// TIA Portal V20 export
// export: Created 2026-10-19T18:06:26.0866612Z, ExportSetting WithDefaults, DisplayName Totally Integrated Automation Portal, DisplayVersion V20 Update 6, DisplayName TIA Portal Openness, DisplayVersion V20 Update 6, DisplayName TIA Portal Version Control Interface, DisplayVersion V20 Update 6, DisplayName SINAMICS Startdrive Advanced, DisplayVersion V20 SP1, DisplayName SINAMICS Startdrive G130, G150, S120, S150, SINAMICS MV, G220, S200, S210, DisplayVersion V20 SP1, DisplayName SINAMICS Startdrive G110M, G120, G120C, G120D, G120P, G115D, DisplayVersion V20 SP1, DisplayName STEP 7 Professional, DisplayVersion V20 Update 6, DisplayName STEP 7 Safety, DisplayVersion V20 Update 2, DisplayName WinCC Basic/Comfort/Advanced, DisplayVersion V20 Update 6, DisplayName WinCC Unified, DisplayVersion V20 Update 6
FUNCTION_BLOCK "SAI_IND_SpanAdjust"   // FB55, LAD
TITLE = Span and Linearity Adjustment (Multi-Point Selectable)
{ S7_Optimized_Access := 'FALSE' }
VERSION : 0.1
// stored: AutoNumber true, IsIECCheckEnabled false, SetENOAutomatically false, UDAEnableTagReadback false
   VAR_INPUT
      ID : HW_IO;   // The Profinet Device Hardware Identifier under device properties
      Hi_Weight : Real;   // The highest adjustment weight, or the Span value
      Mid_Weight : Real;   // The 4th adjustment weight
      Low_Weight : Real;   // The 3rd adjustment weight
      xLow_Weight : Real;   // The 2nd adjustment weight
   END_VAR
   VAR_OUTPUT
      CurrentPoint : Int;   // Current point to be adjusted (Minimum 2 points; maximum 5 points; zero point is the 1st point)
      CurrentWeight : Real;   // Current adjustment weight to be loaded onto the scale
      LoadWeight : Bool;   // Load the next adjustment weight according to value shown in CurrentWeight
      Process : Bool;   // Weight Transmitter is performing adjustment
      Done : Bool;   // Linearity Adjustment has been completed successfully
      Error : Bool;   // Adjustment can not proceed due to incomplete input parameters, check LinearityRange and all the adjustment weight values
      Cancelled : Bool;   // Adjustment process has been cancelled successfully
   END_VAR
   VAR_IN_OUT
      LinearityRange : Int;   // Number of linearity points to be adjusted: 0:none, 1:3 point, 2:4 point, 3:5 point
      Start : Bool;   // Trigger this bit ON to start performing linearity adjustment; this bit will be turned off automatically after completion
      ConfirmWeight : Bool;   // Switch ON this bit as an acknowledgement that new adjustment weight has being loaded
      Cancel : Bool;   // Cancel/ Abort adjustment process, toggle ON
   END_VAR
   VAR DB_SPECIFIC
      Activate : Bool;
   END_VAR
   VAR
      WRREC_SpanAdjust { S7_SetPoint := 'True'} : WRREC;
      RDREC_Status { S7_SetPoint := 'True'} : RDREC;
   END_VAR
   VAR DB_SPECIFIC
      IEC_Timer_1_Instance { S7_SetPoint := 'True'} : IEC_TIMER;
      AdjustStep : SInt;
      Static01 : Bool;
      Static02 : Bool;
      Static03 : Bool;
      Static04 : Bool;
      Static05 : Bool;
      Static06 : Bool;
      Static07 : Bool;
      Static08 : Bool;
      Validate_REC : SInt;
      Abort_REC : SInt;
      Check01 : Bool;
      Check02 : Bool;
      AdjustmentStatus : Int;
      CurrentPoint_0 : Int;
      CurrentWeight_0 : Real;
   END_VAR
   VAR_TEMP   // added for the SCL form of the ladder/FBD networks
      _w1 : Bool;
      _w2 : Bool;
      _w3 : Bool;
      _w4 : Bool;
      _w5 : Bool;
      _w6 : Bool;
      _w7 : Bool;
      _w8 : Bool;
      _w9 : Bool;
      _w10 : Bool;
      _w11 : Bool;
      _w12 : Bool;
      _w13 : Bool;
   END_VAR
BEGIN

REGION Network 1: Initialization
   // Initializes FB output bits:
   // Process;
   // Error;
   // Done;
   // Cancelled
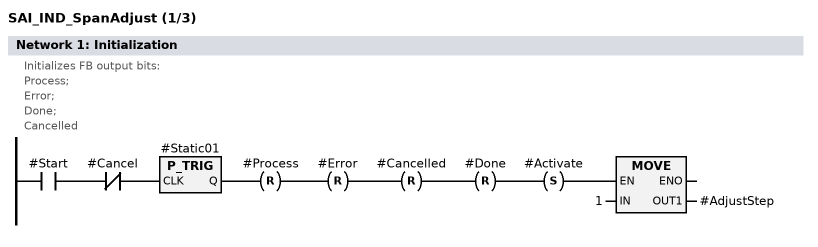
   RUNG wire#powerrail
      Contact( #Start )
      I_Contact( #Cancel )
      P_Trig( #Static01 )
      R_Coil( #Process )
      R_Coil( #Error )
      R_Coil( #Cancelled )
      R_Coil( #Done )
      S_Coil( #Activate )
      { S7_GenerateENO := "TRUE" } Move(in := 1, out1 => #AdjustStep)
   END_RUNG
   // the same network as SCL:
   #_w1 := #Start AND NOT #Cancel;
   #_w2 := #_w1 AND NOT #Static01;   // rising edge
   #Static01 := #_w1;
   IF #_w2 THEN
       #Process := FALSE;
       #Error := FALSE;
       #Cancelled := FALSE;
       #Done := FALSE;
       #Activate := TRUE;
       #AdjustStep := 1;
   END_IF;
END_REGION

REGION Network 2: Sequence
   // AdjustStep = 1: Check all the input parameters for LinearityRange and adjustment weights (Hi_Weight, Mid_Weight, Low_Weight, xLow_Weight)
   // AdjustStep = 2: Initializes all the control bits
   // AdjustStep = 3: Write in the LinearityRange into the transmitter (2-byte; Index: 16#400A)
   // AdjustStep = 4: Updates the CurrentPoint and CurrentWeight (new reference weight) and wait for user to trigger ConfirmWeight input bit
   // AdjustStep = 5: Start the adjustment process according to the CurrentWeight (REAL; Index: 16#4009)
   // AdjustStep = 6: After adjusted all the required reference weights, validate the adjustment (2-byte; Index: 16#4010)
   // AdjustStep = 7: Adjustment is completed successfully, set DONE bit to TRUE
   // AdjustStep = 8; Adjustment failed with error, set ERROR bit to TRUE
   // AdjustStep >= 4: Reading the adjustment status continuously (2-byte; Index: 16#4007)
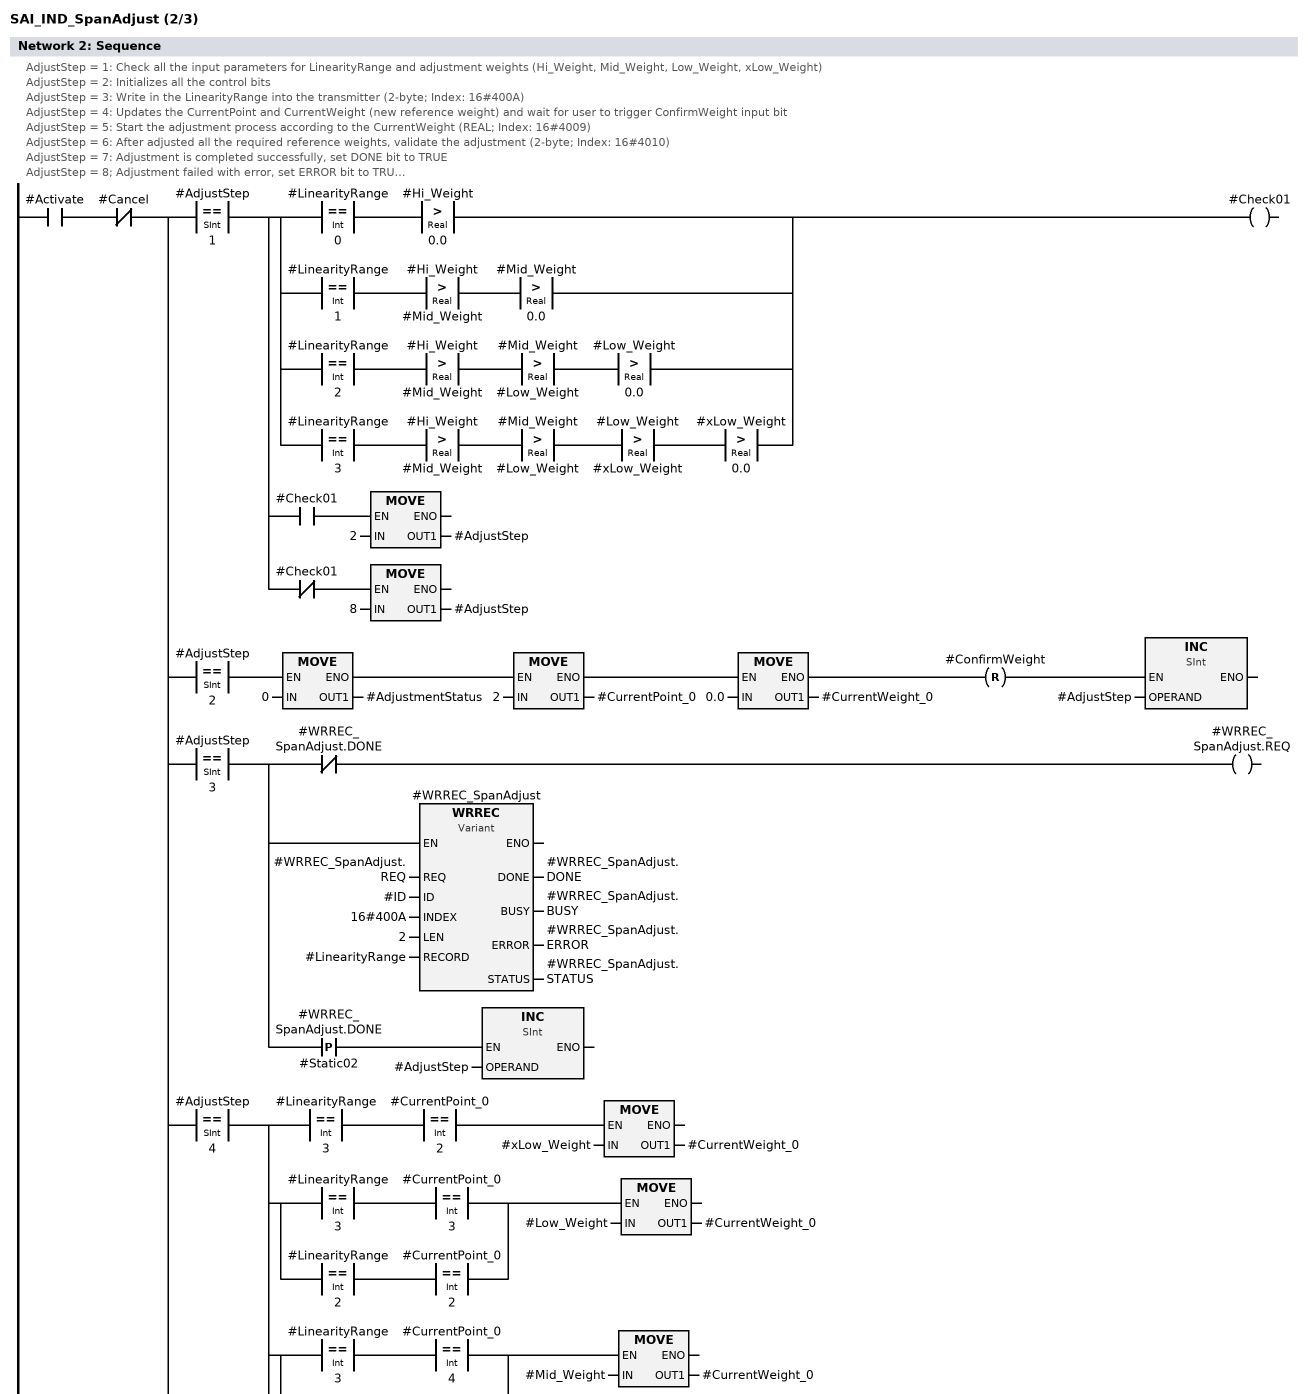
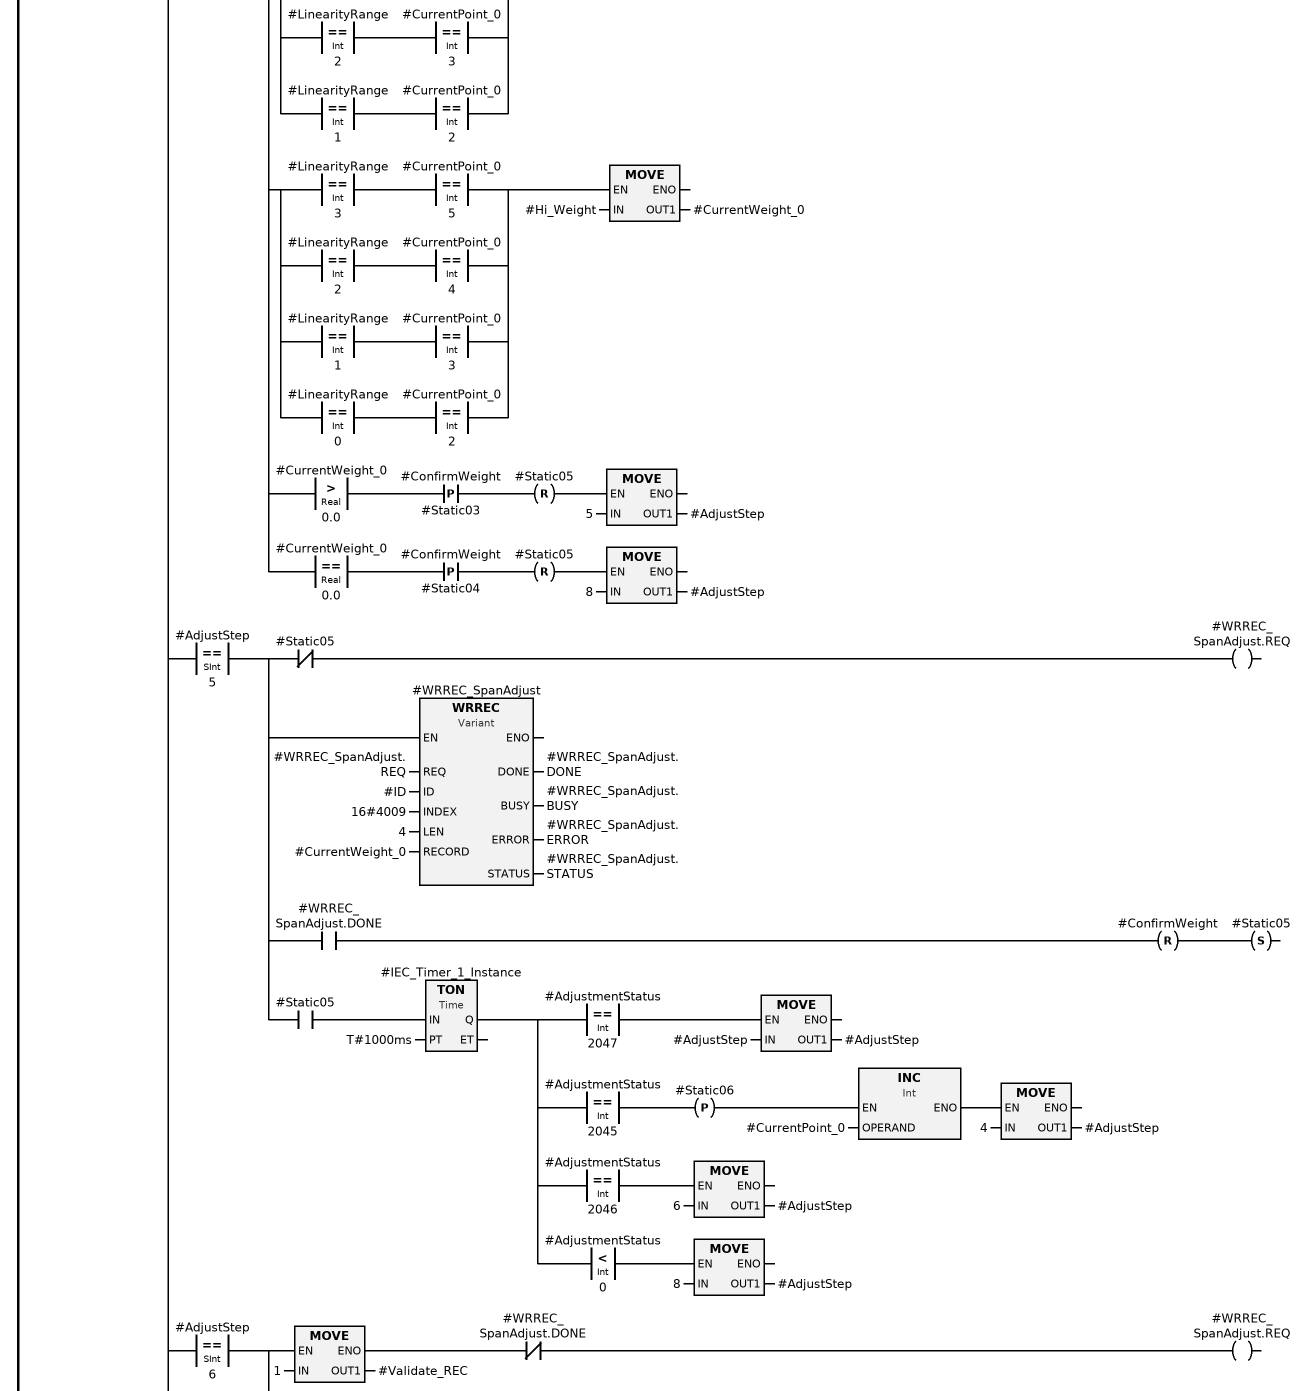
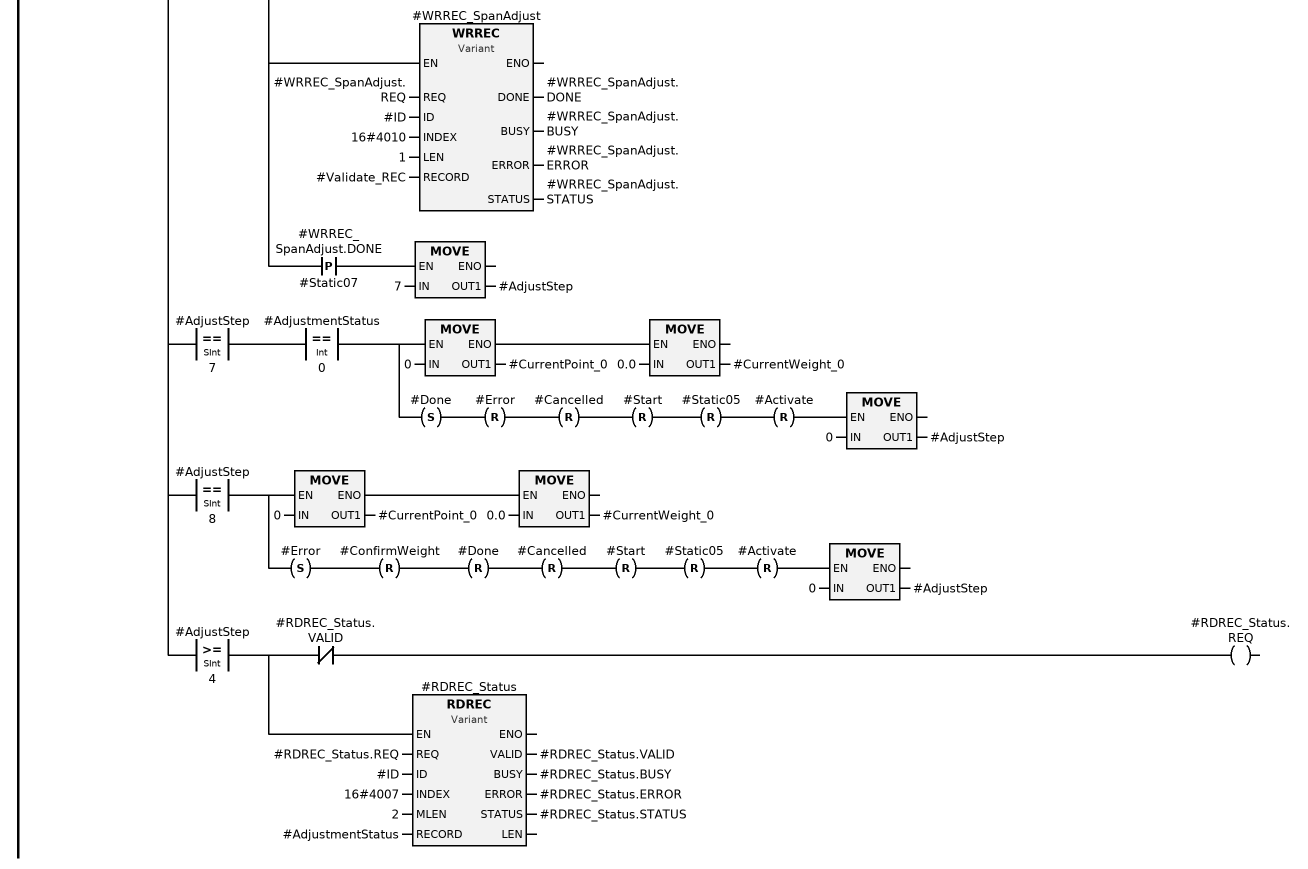
   RUNG wire#powerrail
      Contact( #Activate )
      I_Contact( #Cancel )
      wire#w1
      { S7_Templates := "SrcType := SInt" } EQ_Contact(in1 := #AdjustStep, in2 := 1)
      wire#w2
      { S7_Templates := "SrcType := Int" } EQ_Contact(in1 := #LinearityRange, in2 := 0)
      { S7_Templates := "SrcType := Real" } GT_Contact(in1 := #Hi_Weight, in2 := 0.0)
      wire#w3
      Coil( #Check01 )
   END_RUNG
   RUNG wire#w2
      { S7_Templates := "SrcType := Int" } EQ_Contact(in1 := #LinearityRange, in2 := 1)
      { S7_Templates := "SrcType := Real" } GT_Contact(in1 := #Hi_Weight, in2 := #Mid_Weight)
      { S7_Templates := "SrcType := Real" } GT_Contact(in1 := #Mid_Weight, in2 := 0.0)
   END_RUNG wire#w3
   RUNG wire#w2
      { S7_Templates := "SrcType := Int" } EQ_Contact(in1 := #LinearityRange, in2 := 2)
      { S7_Templates := "SrcType := Real" } GT_Contact(in1 := #Hi_Weight, in2 := #Mid_Weight)
      { S7_Templates := "SrcType := Real" } GT_Contact(in1 := #Mid_Weight, in2 := #Low_Weight)
      { S7_Templates := "SrcType := Real" } GT_Contact(in1 := #Low_Weight, in2 := 0.0)
   END_RUNG wire#w3
   RUNG wire#w2
      { S7_Templates := "SrcType := Int" } EQ_Contact(in1 := #LinearityRange, in2 := 3)
      { S7_Templates := "SrcType := Real" } GT_Contact(in1 := #Hi_Weight, in2 := #Mid_Weight)
      { S7_Templates := "SrcType := Real" } GT_Contact(in1 := #Mid_Weight, in2 := #Low_Weight)
      { S7_Templates := "SrcType := Real" } GT_Contact(in1 := #Low_Weight, in2 := #xLow_Weight)
      { S7_Templates := "SrcType := Real" } GT_Contact(in1 := #xLow_Weight, in2 := 0.0)
   END_RUNG wire#w3
   RUNG wire#w2
      Contact( #Check01 )
      Move(in := 2, out1 => #AdjustStep)
   END_RUNG
   RUNG wire#w2
      I_Contact( #Check01 )
      Move(in := 8, out1 => #AdjustStep)
   END_RUNG
   RUNG wire#w1
      { S7_Templates := "SrcType := SInt" } EQ_Contact(in1 := #AdjustStep, in2 := 2)
      Move(in := 0, out1 => #AdjustmentStatus)
      Move(in := 2, out1 => #CurrentPoint_0)
      Move(in := 0.0, out1 => #CurrentWeight_0)
      R_Coil( #ConfirmWeight )
      { S7_Templates := "DestType := SInt" } Inc( #AdjustStep )
   END_RUNG
   RUNG wire#w1
      { S7_Templates := "SrcType := SInt" } EQ_Contact(in1 := #AdjustStep, in2 := 3)
      wire#w4
      I_Contact( #WRREC_SpanAdjust.DONE )
      Coil( #WRREC_SpanAdjust.REQ )
   END_RUNG
   RUNG wire#w4
      { S7_Templates := "[ptr_type := Variant, id_type := HW_IO, index_type := DInt, len_type := UInt]" } #WRREC_SpanAdjust.WRREC(REQ := #WRREC_SpanAdjust.REQ, ID := #ID, INDEX := 16#400A, LEN := 2, RECORD := #LinearityRange, DONE => #WRREC_SpanAdjust.DONE, BUSY => #WRREC_SpanAdjust.BUSY, ERROR => #WRREC_SpanAdjust.ERROR, STATUS => #WRREC_SpanAdjust.STATUS)
   END_RUNG
   RUNG wire#w4
      P_Contact(operand := #WRREC_SpanAdjust.DONE, bit := #Static02)
      { S7_Templates := "DestType := SInt" } Inc( #AdjustStep )
   END_RUNG
   RUNG wire#w1
      { S7_Templates := "SrcType := SInt" } EQ_Contact(in1 := #AdjustStep, in2 := 4)
      wire#w5
      { S7_Templates := "SrcType := Int" } EQ_Contact(in1 := #LinearityRange, in2 := 3)
      { S7_Templates := "SrcType := Int" } EQ_Contact(in1 := #CurrentPoint_0, in2 := 2)
      Move(in := #xLow_Weight, out1 => #CurrentWeight_0)
   END_RUNG
   RUNG wire#w5
      { S7_Templates := "SrcType := Int" } EQ_Contact(in1 := #LinearityRange, in2 := 3)
      { S7_Templates := "SrcType := Int" } EQ_Contact(in1 := #CurrentPoint_0, in2 := 3)
      wire#w6
      Move(in := #Low_Weight, out1 => #CurrentWeight_0)
   END_RUNG
   RUNG wire#w5
      { S7_Templates := "SrcType := Int" } EQ_Contact(in1 := #LinearityRange, in2 := 2)
      { S7_Templates := "SrcType := Int" } EQ_Contact(in1 := #CurrentPoint_0, in2 := 2)
   END_RUNG wire#w6
   RUNG wire#w5
      { S7_Templates := "SrcType := Int" } EQ_Contact(in1 := #LinearityRange, in2 := 3)
      { S7_Templates := "SrcType := Int" } EQ_Contact(in1 := #CurrentPoint_0, in2 := 4)
      wire#w7
      Move(in := #Mid_Weight, out1 => #CurrentWeight_0)
   END_RUNG
   RUNG wire#w5
      { S7_Templates := "SrcType := Int" } EQ_Contact(in1 := #LinearityRange, in2 := 2)
      { S7_Templates := "SrcType := Int" } EQ_Contact(in1 := #CurrentPoint_0, in2 := 3)
   END_RUNG wire#w7
   RUNG wire#w5
      { S7_Templates := "SrcType := Int" } EQ_Contact(in1 := #LinearityRange, in2 := 1)
      { S7_Templates := "SrcType := Int" } EQ_Contact(in1 := #CurrentPoint_0, in2 := 2)
   END_RUNG wire#w7
   RUNG wire#w5
      { S7_Templates := "SrcType := Int" } EQ_Contact(in1 := #LinearityRange, in2 := 3)
      { S7_Templates := "SrcType := Int" } EQ_Contact(in1 := #CurrentPoint_0, in2 := 5)
      wire#w8
      Move(in := #Hi_Weight, out1 => #CurrentWeight_0)
   END_RUNG
   RUNG wire#w5
      { S7_Templates := "SrcType := Int" } EQ_Contact(in1 := #LinearityRange, in2 := 2)
      { S7_Templates := "SrcType := Int" } EQ_Contact(in1 := #CurrentPoint_0, in2 := 4)
   END_RUNG wire#w8
   RUNG wire#w5
      { S7_Templates := "SrcType := Int" } EQ_Contact(in1 := #LinearityRange, in2 := 1)
      { S7_Templates := "SrcType := Int" } EQ_Contact(in1 := #CurrentPoint_0, in2 := 3)
   END_RUNG wire#w8
   RUNG wire#w5
      { S7_Templates := "SrcType := Int" } EQ_Contact(in1 := #LinearityRange, in2 := 0)
      { S7_Templates := "SrcType := Int" } EQ_Contact(in1 := #CurrentPoint_0, in2 := 2)
   END_RUNG wire#w8
   RUNG wire#w5
      { S7_Templates := "SrcType := Real" } GT_Contact(in1 := #CurrentWeight_0, in2 := 0.0)
      P_Contact(operand := #ConfirmWeight, bit := #Static03)
      R_Coil( #Static05 )
      Move(in := 5, out1 => #AdjustStep)
   END_RUNG
   RUNG wire#w5
      { S7_Templates := "SrcType := Real" } EQ_Contact(in1 := #CurrentWeight_0, in2 := 0.0)
      P_Contact(operand := #ConfirmWeight, bit := #Static04)
      R_Coil( #Static05 )
      Move(in := 8, out1 => #AdjustStep)
   END_RUNG
   RUNG wire#w1
      { S7_Templates := "SrcType := SInt" } EQ_Contact(in1 := #AdjustStep, in2 := 5)
      wire#w9
      I_Contact( #Static05 )
      Coil( #WRREC_SpanAdjust.REQ )
   END_RUNG
   RUNG wire#w9
      { S7_Templates := "[ptr_type := Variant, id_type := HW_IO, index_type := DInt, len_type := UInt]" } #WRREC_SpanAdjust.WRREC(REQ := #WRREC_SpanAdjust.REQ, ID := #ID, INDEX := 16#4009, LEN := 4, RECORD := #CurrentWeight_0, DONE => #WRREC_SpanAdjust.DONE, BUSY => #WRREC_SpanAdjust.BUSY, ERROR => #WRREC_SpanAdjust.ERROR, STATUS => #WRREC_SpanAdjust.STATUS)
   END_RUNG
   RUNG wire#w9
      Contact( #WRREC_SpanAdjust.DONE )
      R_Coil( #ConfirmWeight )
      S_Coil( #Static05 )
   END_RUNG
   RUNG wire#w9
      Contact( #Static05 )
      { S7_Templates := "time_type := Time" } #IEC_Timer_1_Instance.TON(pt := T#1000ms, et =>)
      wire#w10
      { S7_Templates := "SrcType := Int" } EQ_Contact(in1 := #AdjustmentStatus, in2 := 2047)
      Move(in := #AdjustStep, out1 => #AdjustStep)
   END_RUNG
   RUNG wire#w10
      { S7_Templates := "SrcType := Int" } EQ_Contact(in1 := #AdjustmentStatus, in2 := 2045)
      P_Trig( #Static06 )
      { S7_Templates := "DestType := Int" } Inc( #CurrentPoint_0 )
      Move(in := 4, out1 => #AdjustStep)
   END_RUNG
   RUNG wire#w10
      { S7_Templates := "SrcType := Int" } EQ_Contact(in1 := #AdjustmentStatus, in2 := 2046)
      Move(in := 6, out1 => #AdjustStep)
   END_RUNG
   RUNG wire#w10
      { S7_Templates := "SrcType := Int" } LT_Contact(in1 := #AdjustmentStatus, in2 := 0)
      Move(in := 8, out1 => #AdjustStep)
   END_RUNG
   RUNG wire#w1
      { S7_Templates := "SrcType := SInt" } EQ_Contact(in1 := #AdjustStep, in2 := 6)
      wire#w11
      Move(in := 1, out1 => #Validate_REC)
      I_Contact( #WRREC_SpanAdjust.DONE )
      Coil( #WRREC_SpanAdjust.REQ )
   END_RUNG
   RUNG wire#w11
      { S7_Templates := "[ptr_type := Variant, id_type := HW_IO, index_type := DInt, len_type := UInt]" } #WRREC_SpanAdjust.WRREC(REQ := #WRREC_SpanAdjust.REQ, ID := #ID, INDEX := 16#4010, LEN := 1, RECORD := #Validate_REC, DONE => #WRREC_SpanAdjust.DONE, BUSY => #WRREC_SpanAdjust.BUSY, ERROR => #WRREC_SpanAdjust.ERROR, STATUS => #WRREC_SpanAdjust.STATUS)
   END_RUNG
   RUNG wire#w11
      P_Contact(operand := #WRREC_SpanAdjust.DONE, bit := #Static07)
      Move(in := 7, out1 => #AdjustStep)
   END_RUNG
   RUNG wire#w1
      { S7_Templates := "SrcType := SInt" } EQ_Contact(in1 := #AdjustStep, in2 := 7)
      { S7_Templates := "SrcType := Int" } EQ_Contact(in1 := #AdjustmentStatus, in2 := 0)
      wire#w12
      Move(in := 0, out1 => #CurrentPoint_0)
      Move(in := 0.0, out1 => #CurrentWeight_0)
   END_RUNG
   RUNG wire#w12
      S_Coil( #Done )
      R_Coil( #Error )
      R_Coil( #Cancelled )
      R_Coil( #Start )
      R_Coil( #Static05 )
      R_Coil( #Activate )
      Move(in := 0, out1 => #AdjustStep)
   END_RUNG
   RUNG wire#w1
      { S7_Templates := "SrcType := SInt" } EQ_Contact(in1 := #AdjustStep, in2 := 8)
      wire#w13
      Move(in := 0, out1 => #CurrentPoint_0)
      Move(in := 0.0, out1 => #CurrentWeight_0)
   END_RUNG
   RUNG wire#w13
      S_Coil( #Error )
      R_Coil( #ConfirmWeight )
      R_Coil( #Done )
      R_Coil( #Cancelled )
      R_Coil( #Start )
      R_Coil( #Static05 )
      R_Coil( #Activate )
      Move(in := 0, out1 => #AdjustStep)
   END_RUNG
   RUNG wire#w1
      { S7_Templates := "SrcType := SInt" } GE_Contact(in1 := #AdjustStep, in2 := 4)
      wire#w14
      I_Contact( #RDREC_Status.VALID )
      Coil( #RDREC_Status.REQ )
   END_RUNG
   RUNG wire#w14
      { S7_Templates := "[ptr_type := Variant, id_type := HW_IO, index_type := DInt, len_type := UInt]" } #RDREC_Status.RDREC(REQ := #RDREC_Status.REQ, ID := #ID, INDEX := 16#4007, MLEN := 2, RECORD := #AdjustmentStatus, VALID => #RDREC_Status.VALID, BUSY => #RDREC_Status.BUSY, ERROR => #RDREC_Status.ERROR, STATUS => #RDREC_Status.STATUS, LEN =>)
   END_RUNG
   // the same network as SCL:
   #_w1 := #Activate AND NOT #Cancel;
   #_w2 := #_w1 AND (#AdjustStep = 1);
   #Check01 := #_w2 AND (((#LinearityRange = 0) AND (#Hi_Weight > 0.0)) OR ((#LinearityRange = 1) AND (#Hi_Weight > #Mid_Weight) AND (#Mid_Weight > 0.0)) OR ((#LinearityRange = 2) AND (#Hi_Weight > #Mid_Weight) AND (#Mid_Weight > #Low_Weight) AND (#Low_Weight > 0.0)) OR ((#LinearityRange = 3) AND (#Hi_Weight > #Mid_Weight) AND (#Mid_Weight > #Low_Weight) AND (#Low_Weight > #xLow_Weight) AND (#xLow_Weight > 0.0)));
   IF #_w2 AND #Check01 THEN #AdjustStep := 2; END_IF;
   IF #_w2 AND NOT #Check01 THEN #AdjustStep := 8; END_IF;
   IF #_w1 AND (#AdjustStep = 2) THEN
       #AdjustmentStatus := 0;
       #CurrentPoint_0 := 2;
       #CurrentWeight_0 := 0.0;
       #ConfirmWeight := FALSE;
       #AdjustStep := #AdjustStep + 1;
   END_IF;
   #_w3 := #_w1 AND (#AdjustStep = 3);
   #WRREC_SpanAdjust.REQ := #_w3 AND NOT #WRREC_SpanAdjust.DONE;
   IF #_w3 THEN
       #WRREC_SpanAdjust(REQ := #WRREC_SpanAdjust.REQ,   // WRREC
                         ID := #ID,
                         INDEX := 16#400A,
                         LEN := 2,
                         RECORD := #LinearityRange,
                         DONE => #WRREC_SpanAdjust.DONE,
                         BUSY => #WRREC_SpanAdjust.BUSY,
                         ERROR => #WRREC_SpanAdjust.ERROR,
                         STATUS => #WRREC_SpanAdjust.STATUS);
   END_IF;
   #_w4 := #_w3 AND #WRREC_SpanAdjust.DONE AND NOT #Static02;   // rising edge of #WRREC_SpanAdjust.DONE
   #Static02 := #WRREC_SpanAdjust.DONE;
   IF #_w4 THEN #AdjustStep := #AdjustStep + 1; END_IF;
   #_w5 := #_w1 AND (#AdjustStep = 4);
   IF #_w5 AND (#LinearityRange = 3) AND (#CurrentPoint_0 = 2) THEN #CurrentWeight_0 := #xLow_Weight; END_IF;
   IF #_w5 AND (((#LinearityRange = 3) AND (#CurrentPoint_0 = 3)) OR ((#LinearityRange = 2) AND (#CurrentPoint_0 = 2))) THEN
       #CurrentWeight_0 := #Low_Weight;
   END_IF;
   IF #_w5 AND (((#LinearityRange = 3) AND (#CurrentPoint_0 = 4)) OR ((#LinearityRange = 2) AND (#CurrentPoint_0 = 3)) OR ((#LinearityRange = 1) AND (#CurrentPoint_0 = 2))) THEN
       #CurrentWeight_0 := #Mid_Weight;
   END_IF;
   IF #_w5 AND (((#LinearityRange = 3) AND (#CurrentPoint_0 = 5)) OR ((#LinearityRange = 2) AND (#CurrentPoint_0 = 4)) OR ((#LinearityRange = 1) AND (#CurrentPoint_0 = 3)) OR ((#LinearityRange = 0) AND (#CurrentPoint_0 = 2))) THEN
       #CurrentWeight_0 := #Hi_Weight;
   END_IF;
   #_w6 := #_w5 AND (#CurrentWeight_0 > 0.0) AND #ConfirmWeight AND NOT #Static03;   // rising edge of #ConfirmWeight
   #Static03 := #ConfirmWeight;
   IF #_w6 THEN
       #Static05 := FALSE;
       #AdjustStep := 5;
   END_IF;
   #_w7 := #_w5 AND (#CurrentWeight_0 = 0.0) AND #ConfirmWeight AND NOT #Static04;   // rising edge of #ConfirmWeight
   #Static04 := #ConfirmWeight;
   IF #_w7 THEN
       #Static05 := FALSE;
       #AdjustStep := 8;
   END_IF;
   #_w8 := #_w1 AND (#AdjustStep = 5);
   #WRREC_SpanAdjust.REQ := #_w8 AND NOT #Static05;
   IF #_w8 THEN
       #WRREC_SpanAdjust(REQ := #WRREC_SpanAdjust.REQ,   // WRREC
                         ID := #ID,
                         INDEX := 16#4009,
                         LEN := 4,
                         RECORD := #CurrentWeight_0,
                         DONE => #WRREC_SpanAdjust.DONE,
                         BUSY => #WRREC_SpanAdjust.BUSY,
                         ERROR => #WRREC_SpanAdjust.ERROR,
                         STATUS => #WRREC_SpanAdjust.STATUS);
   END_IF;
   IF #_w8 AND #WRREC_SpanAdjust.DONE THEN
       #ConfirmWeight := FALSE;
       #Static05 := TRUE;
   END_IF;
   #IEC_Timer_1_Instance.TON(IN := #_w8 AND #Static05, PT := T#1000ms);
   IF #IEC_Timer_1_Instance.Q AND (#AdjustmentStatus = 2047) THEN #AdjustStep := #AdjustStep; END_IF;
   #_w9 := #IEC_Timer_1_Instance.Q AND (#AdjustmentStatus = 2045);
   #_w10 := #_w9 AND NOT #Static06;   // rising edge
   #Static06 := #_w9;
   IF #_w10 THEN
       #CurrentPoint_0 := #CurrentPoint_0 + 1;
       #AdjustStep := 4;
   END_IF;
   IF #IEC_Timer_1_Instance.Q AND (#AdjustmentStatus = 2046) THEN #AdjustStep := 6; END_IF;
   IF #IEC_Timer_1_Instance.Q AND (#AdjustmentStatus < 0) THEN #AdjustStep := 8; END_IF;
   #_w11 := #_w1 AND (#AdjustStep = 6);
   IF #_w11 THEN #Validate_REC := 1; END_IF;
   #WRREC_SpanAdjust.REQ := #_w11 AND NOT #WRREC_SpanAdjust.DONE;
   IF #_w11 THEN
       #WRREC_SpanAdjust(REQ := #WRREC_SpanAdjust.REQ,   // WRREC
                         ID := #ID,
                         INDEX := 16#4010,
                         LEN := 1,
                         RECORD := #Validate_REC,
                         DONE => #WRREC_SpanAdjust.DONE,
                         BUSY => #WRREC_SpanAdjust.BUSY,
                         ERROR => #WRREC_SpanAdjust.ERROR,
                         STATUS => #WRREC_SpanAdjust.STATUS);
   END_IF;
   #_w12 := #_w11 AND #WRREC_SpanAdjust.DONE AND NOT #Static07;   // rising edge of #WRREC_SpanAdjust.DONE
   #Static07 := #WRREC_SpanAdjust.DONE;
   IF #_w12 THEN #AdjustStep := 7; END_IF;
   IF #_w1 AND (#AdjustStep = 7) AND (#AdjustmentStatus = 0) THEN
       #CurrentPoint_0 := 0;
       #CurrentWeight_0 := 0.0;
       #Done := TRUE;
       #Error := FALSE;
       #Cancelled := FALSE;
       #Start := FALSE;
       #Static05 := FALSE;
       #Activate := FALSE;
       #AdjustStep := 0;
   END_IF;
   IF #_w1 AND (#AdjustStep = 8) THEN
       #CurrentPoint_0 := 0;
       #CurrentWeight_0 := 0.0;
       #Error := TRUE;
       #ConfirmWeight := FALSE;
       #Done := FALSE;
       #Cancelled := FALSE;
       #Start := FALSE;
       #Static05 := FALSE;
       #Activate := FALSE;
       #AdjustStep := 0;
   END_IF;
   #_w13 := #_w1 AND (#AdjustStep >= 4);
   #RDREC_Status.REQ := #_w13 AND NOT #RDREC_Status.VALID;
   IF #_w13 THEN
       #RDREC_Status(REQ := #RDREC_Status.REQ,   // RDREC
                     ID := #ID,
                     INDEX := 16#4007,
                     MLEN := 2,
                     RECORD := #AdjustmentStatus,
                     VALID => #RDREC_Status.VALID,
                     BUSY => #RDREC_Status.BUSY,
                     ERROR => #RDREC_Status.ERROR,
                     STATUS => #RDREC_Status.STATUS);
   END_IF;
END_REGION

REGION Network 3: Adjsutment Status
   // LoadWeight - Inform user to load the next adjustment weight according to CurrentWeight value
   // Process - Status bit to inform that the weight transmitter is performing adjustment process
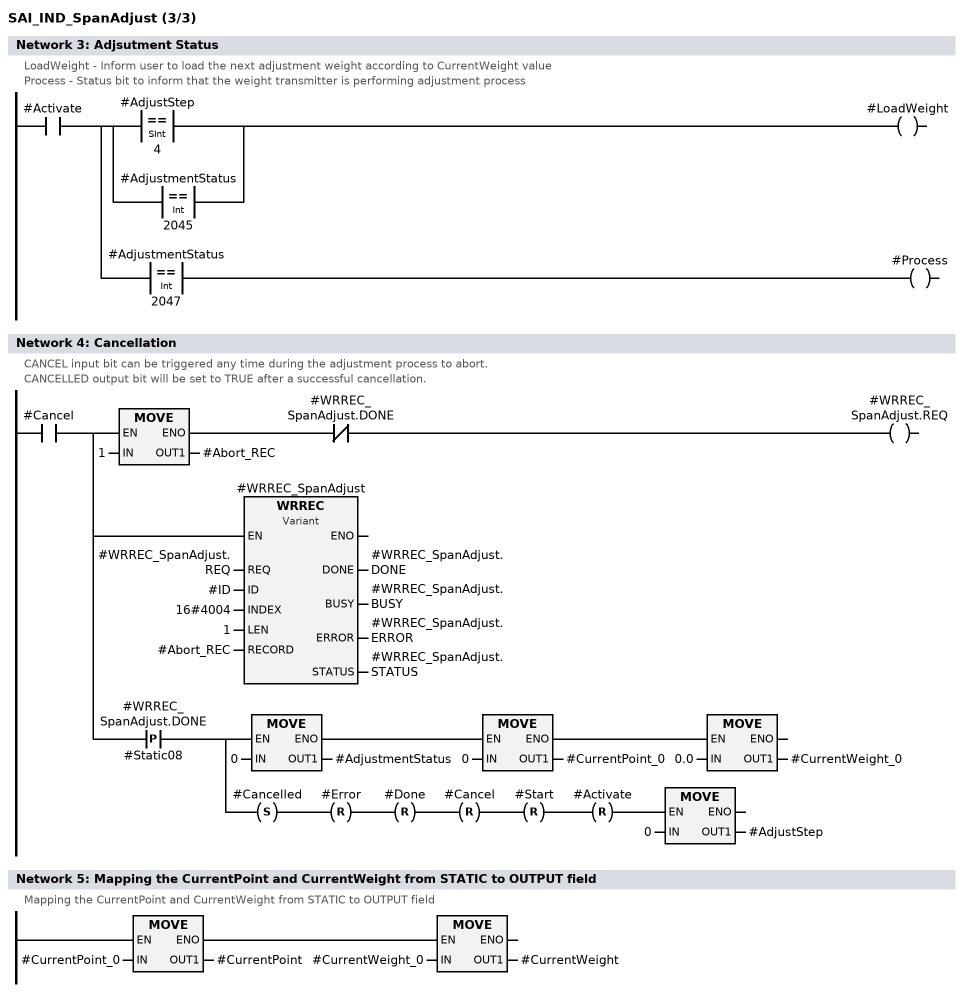
   RUNG wire#powerrail
      Contact( #Activate )
      wire#w1
      { S7_Templates := "SrcType := SInt" } EQ_Contact(in1 := #AdjustStep, in2 := 4)
      wire#w2
      Coil( #LoadWeight )
   END_RUNG
   RUNG wire#w1
      { S7_Templates := "SrcType := Int" } EQ_Contact(in1 := #AdjustmentStatus, in2 := 2045)
   END_RUNG wire#w2
   RUNG wire#w1
      { S7_Templates := "SrcType := Int" } EQ_Contact(in1 := #AdjustmentStatus, in2 := 2047)
      Coil( #Process )
   END_RUNG
   // the same network as SCL:
   #LoadWeight := #Activate AND ((#AdjustStep = 4) OR (#AdjustmentStatus = 2045));
   #Process := #Activate AND (#AdjustmentStatus = 2047);
END_REGION

REGION Network 4: Cancellation
   // CANCEL input bit can be triggered any time during the adjustment process to abort. 
   // CANCELLED output bit will be set to TRUE after a successful cancellation.
   RUNG wire#powerrail
      Contact( #Cancel )
      wire#w1
      Move(in := 1, out1 => #Abort_REC)
      I_Contact( #WRREC_SpanAdjust.DONE )
      Coil( #WRREC_SpanAdjust.REQ )
   END_RUNG
   RUNG wire#w1
      { S7_Templates := "[ptr_type := Variant, id_type := HW_IO, index_type := DInt, len_type := UInt]" } #WRREC_SpanAdjust.WRREC(REQ := #WRREC_SpanAdjust.REQ, ID := #ID, INDEX := 16#4004, LEN := 1, RECORD := #Abort_REC, DONE => #WRREC_SpanAdjust.DONE, BUSY => #WRREC_SpanAdjust.BUSY, ERROR => #WRREC_SpanAdjust.ERROR, STATUS => #WRREC_SpanAdjust.STATUS)
   END_RUNG
   RUNG wire#w1
      P_Contact(operand := #WRREC_SpanAdjust.DONE, bit := #Static08)
      wire#w2
      Move(in := 0, out1 => #AdjustmentStatus)
      Move(in := 0, out1 => #CurrentPoint_0)
      Move(in := 0.0, out1 => #CurrentWeight_0)
   END_RUNG
   RUNG wire#w2
      S_Coil( #Cancelled )
      R_Coil( #Error )
      R_Coil( #Done )
      R_Coil( #Cancel )
      R_Coil( #Start )
      R_Coil( #Activate )
      Move(in := 0, out1 => #AdjustStep)
   END_RUNG
   // the same network as SCL:
   IF #Cancel THEN #Abort_REC := 1; END_IF;
   #WRREC_SpanAdjust.REQ := #Cancel AND NOT #WRREC_SpanAdjust.DONE;
   IF #Cancel THEN
       #WRREC_SpanAdjust(REQ := #WRREC_SpanAdjust.REQ,   // WRREC
                         ID := #ID,
                         INDEX := 16#4004,
                         LEN := 1,
                         RECORD := #Abort_REC,
                         DONE => #WRREC_SpanAdjust.DONE,
                         BUSY => #WRREC_SpanAdjust.BUSY,
                         ERROR => #WRREC_SpanAdjust.ERROR,
                         STATUS => #WRREC_SpanAdjust.STATUS);
   END_IF;
   #_w1 := #Cancel AND #WRREC_SpanAdjust.DONE AND NOT #Static08;   // rising edge of #WRREC_SpanAdjust.DONE
   #Static08 := #WRREC_SpanAdjust.DONE;
   IF #_w1 THEN
       #AdjustmentStatus := 0;
       #CurrentPoint_0 := 0;
       #CurrentWeight_0 := 0.0;
       #Cancelled := TRUE;
       #Error := FALSE;
       #Done := FALSE;
       #Cancel := FALSE;
       #Start := FALSE;
       #Activate := FALSE;
       #AdjustStep := 0;
   END_IF;
END_REGION

REGION Network 5: Mapping the CurrentPoint and CurrentWeight from STATIC to OUTPUT field
   // Mapping the CurrentPoint and CurrentWeight from STATIC to OUTPUT field
   RUNG wire#powerrail
      Move(in := #CurrentPoint_0, out1 => #CurrentPoint)
      Move(in := #CurrentWeight_0, out1 => #CurrentWeight)
   END_RUNG
   // the same network as SCL:
   #CurrentPoint := #CurrentPoint_0;
   #CurrentWeight := #CurrentWeight_0;
END_REGION
END_FUNCTION_BLOCK
